// TIA Portal V21 export
// export: Created 2026-10-23T20:42:08.4059799Z, ExportSetting WithDefaults, DisplayName Totally Integrated Automation Portal, DisplayVersion V21 Update 1, DisplayName SINAMICS Startdrive Advanced, DisplayVersion V21 HF2, DisplayName SINAMICS Startdrive G110M, G120, G120C, G120D, G120P, G115D, DisplayVersion V21 HF2, DisplayName SINAMICS Startdrive G130, G150, S120, S150, G200, G220, S200, S210, S220, Innomotics MVD, DisplayVersion V21 HF2, DisplayName STEP 7 Professional, DisplayVersion V21 Update 1, DisplayName STEP 7 Safety, DisplayVersion V21, DisplayName Tech WebApplication, DisplayVersion V21, DisplayName WinCC Basic/Comfort/Advanced, DisplayVersion V21 Update 1, DisplayName WinCC Unified, DisplayVersion V21 Update 1
ORGANIZATION_BLOCK "OB_Startup"   // OB100, SCL, Startup
TITLE = Anlauf / Startup
{ S7_Optimized_Access := 'TRUE' }
VERSION : 0.1
// Initialisiert Maschinendaten beim Anlauf / Initialises machine data at startup
// stored: AutoNumber false, IsIECCheckEnabled false, SetENOAutomatically false
   VAR_INPUT
      LostRetentive : Bool;   // True if retentive data are lost
      LostRTC : Bool;   // True if date and time are lost
   END_VAR
BEGIN

       REGION Initialise machine data
           "DB_Machine".MachineOn := FALSE;
           "DB_Machine".PieceCount := 0;
           "DB_Machine".SpeedSetpoint := 50.0;
           "DB_Machine".MachineName := 'Filler';
       END_REGION
END_ORGANIZATION_BLOCK
